(* IEC 61131-3 sources: nautilus/website/lessons/b1-blink/start, 1 file *)

(* ---- program.st ---- *)
PROGRAM Blink
VAR
    tick : TON;   (* a half-second stopwatch *)
END_VAR

(* TODO 1: start the stopwatch, and restart it each time it finishes. *)

(* TODO 2: when the stopwatch finishes, flip Lamp. *)

END_PROGRAM
